(* IEC 61131-3 sources: 2026_Projet_YGO_ExcavatriceDragage/ARCHIVES/Code/SUPERVISION/_TYPES, 5 files *)

(* ---- ST_InputsQualified.st ---- *)
(* ═══════════════════════════════════════════════════════════════
   🏗️ ST_InputsQualified — TOR réelles qualifiées (squelette 22 entrées)
   ───────────────────────────────────────────────────────────────
   📄 Lot M1 · Doc : DOC/AF_Partie-06_Acquisition_Qualification_IO_v2.1.md §2ter/§4
   🎨 Une entrée BOOL par TOR réelle qualifiée, organisée par domaine
      (Winch 8 · Translation 7 · Machine 7 = 22).
   🔗 Producteur : PRG_01_Inputs_LD (Ladder, FB_Input) — écrivain unique.
      Lecteur : PRG_02_Acquisition_CFC (seul — alimente le « réel » des domaines TOR).
   ✅ Polarité : TRUE = état logique normalisé (déjà inversé/filtré par FB_Input).
      Filtre appliqué avant la sélection, sur le réel uniquement (décision Q1=A).
      Aucune simulation n'y figure : la bascule réel/simulé vit dans PRG_02.
   ═══════════════════════════════════════════════════════════════ *)
TYPE ST_InputsQualified :
STRUCT
    Winch       : ST_InputsQualifiedWinch;       (* TOR réelles qualifiées Treuils M1/M2 *)
    Translation : ST_InputsQualifiedTranslation; (* TOR réelles qualifiées Translation M3 *)
    Machine     : ST_InputsQualifiedMachine;     (* TOR réelles qualifiées Sécurités/Communs *)
END_STRUCT
END_TYPE

(* ---- ST_InputsQualifiedMachine.st ---- *)
(* ═══════════════════════════════════════════════════════════════
   🏗️ ST_InputsQualifiedMachine — TOR réelles qualifiées domaine Machine
   ───────────────────────────────────────────────────────────────
   📄 Lot M1 (PRG_01_Inputs_LD → ST_InputsQualified)
   🎨 Champs qualifiés (polarité normalisée, filtre FB_Input appliqué).
   🔗 Producteur : PRG_01_Inputs_LD · Lecteur : PRG_02_Acquisition_CFC
   ═══════════════════════════════════════════════════════════════ *)
TYPE ST_InputsQualifiedMachine :
STRUCT
    PowerContactorEngaged_DI   : BOOL; (* TRUE = contacteur de puissance engagé *)
    EmergencyChainClosed_DI    : BOOL; (* TRUE = boucle AU fermée (saine) *)
    PhaseRotationOk_DI         : BOOL; (* TRUE = rotation des phases correcte *)
    BrakeThermalOk_DI          : BOOL; (* TRUE = thermique freins M1/M2/M3 commun OK *)
    M1_M2_KoboldContactFond_DI : BOOL; (* TRUE = contact fond Kobold détecté *)
    HydraulicThermalOk_DI      : BOOL; (* TRUE = thermique moteur hydraulique OK *)
    ConveyorInfeedReady_DI     : BOOL; (* TRUE = autorisation démarrage crible *)
END_STRUCT
END_TYPE

(* ---- ST_InputsQualifiedTranslation.st ---- *)
(* ═══════════════════════════════════════════════════════════════
   🏗️ ST_InputsQualifiedTranslation — TOR réelles qualifiées domaine Translation
   ───────────────────────────────────────────────────────────────
   📄 Lot M1 (PRG_01_Inputs_LD → ST_InputsQualified)
   🎨 Champs qualifiés (polarité normalisée, filtre FB_Input appliqué).
   🔗 Producteur : PRG_01_Inputs_LD · Lecteur : PRG_02_Acquisition_CFC
   ═══════════════════════════════════════════════════════════════ *)
TYPE ST_InputsQualifiedTranslation :
STRUCT
    M3_BrakeIsOpen_DI        : BOOL; (* TRUE = frein M3 OUVERT (desserré) — REX 08-03 *)
    M3_ThermalFeedback_DI    : BOOL; (* TRUE = thermique M3 OK *)
    M3_PosTremie_DI          : BOOL; (* TRUE = chariot en position Trémie *)
    M3_PosPV_DI              : BOOL; (* TRUE = chariot en zone pré-ralentissement PV *)
    M3_PosP2_DI              : BOOL; (* TRUE = chariot en position P2 *)
    M3_PosP1_DI              : BOOL; (* TRUE = chariot en position P1 *)
    M3_PosMaintenance_DI     : BOOL; (* TRUE = chariot en position Maintenance *)
END_STRUCT
END_TYPE

(* ---- ST_InputsQualifiedWinch.st ---- *)
(* ═══════════════════════════════════════════════════════════════
   🏗️ ST_InputsQualifiedWinch — TOR réelles qualifiées domaine Treuils
   ───────────────────────────────────────────────────────────────
   📄 Lot M1 (PRG_01_Inputs_LD → ST_InputsQualified)
   🎨 Champs qualifiés (polarité normalisée, filtre FB_Input appliqué).
   🔗 Producteur : PRG_01_Inputs_LD · Lecteur : PRG_02_Acquisition_CFC
   ═══════════════════════════════════════════════════════════════ *)
TYPE ST_InputsQualifiedWinch :
STRUCT
    M1_ContactorsReleased_DI : BOOL; (* TRUE = contacteurs M1 retombés (sain) *)
    M1_ThermalOk_DI          : BOOL; (* TRUE = thermique M1 OK *)
    M1_BrakeIsOpen_DI        : BOOL; (* TRUE = frein M1 OUVERT (desserré) — REX 08-03 *)
    M2_ContactorsReleased_DI : BOOL; (* TRUE = contacteurs M2 retombés (sain) *)
    M2_ThermalOk_DI          : BOOL; (* TRUE = thermique M2 OK *)
    M2_BrakeIsOpen_DI        : BOOL; (* TRUE = frein M2 OUVERT (desserré) — REX 08-03 *)
    M1M2_TopPositionFree_DI  : BOOL; (* TRUE = fin de course haut libre *)
    M2_TensionedCable_DI     : BOOL; (* TRUE = câble M2 tendu (mou non déclenché) *)
END_STRUCT
END_TYPE

(* ---- ST_OperatorAction.st ---- *)
(* ═══════════════════════════════════════════════════════════════
   🎮 ST_OperatorAction — Consigne unique de conduite opérateur
   ───────────────────────────────────────────────────────────────
   📄 Doc : DOC/AF/AF_Partie-07_Interface_IHM_v2.1.md
   🎯 Les alarmes restent dans Error/ErrorId : cette struct répond seulement
      à « quelle action attend-on maintenant de l'opérateur ? ».
   ═══════════════════════════════════════════════════════════════ *)
TYPE ST_OperatorAction :
STRUCT
    ActionId : WORD;        (* Identifiant stable : table de textes IHM possible *)
    Text     : STRING(120); (* Texte de secours pour IHM/diagnostic acceptant les STRING *)
END_STRUCT
END_TYPE
